Fanuc KAREL source: kd00034.KL

-- PROVISIONAL review KL for V940-1; original PC SHA256 19e1e94f56aff58c86a74c9cfccfc9e311d6df2a3dc4bb94dc210021ce49fc8e
-- Incomplete behavior may be omitted. Consult companion uncertainty JSON. Do not deploy.
PROGRAM KD00034
%NOLOCKGROUP
VAR
  I : INTEGER
  J : INTEGER
  B : BOOLEAN
  R : REAL
  S : STRING[80]
BEGIN
  -- V9_ZERO_TABLE_METADATA_HINT layout=0001; no indexed target words; source/name/runtime held
  -- UNRESOLVED_PC offsets 5-27; opcodes 9D,81,18,22,9D,12,22,9D,13,04
  -- UNRESOLVED_PC offsets 32-36; opcodes 7F
END KD00034
